TYPE "ST_SatelliteUnitHal"
VERSION : 0.1
   STRUCT
      "Cell" {ExternalAccessible := 'False'; ExternalVisible := 'False'; ExternalWritable := 'False'} : "ST_DeclarationCellHal";
      "Inner" {ExternalAccessible := 'False'; ExternalVisible := 'False'; ExternalWritable := 'False'} : "ST_InnerUnitHal";
   END_STRUCT;
END_TYPE
